(* IEC 61131-3 sources: codesys-ai-industrial-robot-control/plc/src/Tests, 11 files *)

(* ---- PRG_TestAlarms.st ---- *)
(*
    PRG_TestAlarms
    Purpose : Simulation test harness for FB_AlarmHandler (tests/plc/alarms.json).
    Inputs  : eId + xRaise / xRaiseEvent / xClear pulses, xAck, xReinit (each pulse resets itself).
*)
PROGRAM PRG_TestAlarms
VAR
    fbAlarms : FB_AlarmHandler;
    fbAlarmsInitial : FB_AlarmHandler;
    eId : E_AlarmId;
    xRaise : BOOL;
    xRaiseEvent : BOOL;
    xClear : BOOL;
    xAck : BOOL;
    xReinit : BOOL;
END_VAR

IF xReinit THEN
    xReinit := FALSE;
    fbAlarms := fbAlarmsInitial;
END_IF
IF xRaise THEN
    xRaise := FALSE;
    fbAlarms.Raise(eId);
END_IF
IF xRaiseEvent THEN
    xRaiseEvent := FALSE;
    fbAlarms.RaiseEvent(eId);
END_IF
IF xClear THEN
    xClear := FALSE;
    fbAlarms.Clear(eId);
END_IF
IF xAck THEN
    xAck := FALSE;
    fbAlarms.AcknowledgeAll();
END_IF
fbAlarms();

(* ---- PRG_TestCell.st ---- *)
(*
    PRG_TestCell
    Purpose : Simulation test harness for the whole cell in PRG_Main (tests/plc/cell.json).
              Simulates the vacuum switch, injects parts (PE1 pulse, then vision and decision
              messages for the captured part id) and can press the E-stop or lose the vacuum
              during a transfer. Can play the twin's bridge (heartbeat, joint feedback answering
              the current setpoint sample, twin active) and stall it. While active it plays an AI
              decision service (GVL_Bridge.xDecisionActive), reset when it is switched off.
    Inputs  : xActive; xInject (+ usiInjClass, eInjQuality); xEStopOnTransfer; xVacLostOnTransfer;
              xMark (J1 reference); xBridgeSim; xBridgeStall (heartbeat stops toggling);
              xBridgeStallOnTransfer
    Outputs : lrJ1Delta - J1 movement since xMark [deg]; lrAbortDelayMs - bridge stall -> Aborted
*)
PROGRAM PRG_TestCell
VAR
    xActive : BOOL;
    xWasActive : BOOL;
    xInject : BOOL;
    usiInjClass : USINT;
    eInjQuality : E_Quality := E_Quality.Ok;
    iInject : INT;
    tonPulse : TON;
    tonVac : TON;
    xEStopOnTransfer : BOOL;
    xVacLostOnTransfer : BOOL;
    xVacLost : BOOL;                    // latched until xVacLostOnTransfer is released
    xMark : BOOL;
    lrJ1Start : LREAL;
    lrJ1Delta : LREAL;
    xBridgeSim : BOOL;
    xBridgeStall : BOOL;
    xBridgeStallOnTransfer : BOOL;      // stall the bridge when the robot carries a part to its bin
    xStallTimed : BOOL;
    tStall : TIME;
    lrAbortDelayMs : LREAL;             // stall -> Aborted [ms]
END_VAR
VAR CONSTANT
    PE1_PULSE : TIME := T#250MS;
END_VAR

IF NOT xActive THEN
    IF xWasActive THEN                   // leave no fake decision service behind
        GVL_Bridge.xDecisionActive := FALSE;
        xWasActive := FALSE;
    END_IF
    RETURN;
END_IF
xWasActive := TRUE;
GVL_Bridge.xDecisionActive := TRUE;  // the harness injects AI decisions (eInjQuality)

IF xVacLostOnTransfer AND PRG_Main.fbCell.ePickStep = E_PickStep.MoveToBin THEN
    xVacLost := TRUE;
ELSIF NOT xVacLostOnTransfer THEN
    xVacLost := FALSE;
END_IF
tonVac(IN := GVL_Bridge.xVacuumOn, PT := T#100MS);
GVL_Bridge.xVacuumOk := tonVac.Q AND NOT xVacLost;

// the twin's bridge: feedback answers the current setpoint sample, heartbeat toggles
IF xBridgeStallOnTransfer AND NOT xBridgeStall AND PRG_Main.fbCell.ePickStep = E_PickStep.MoveToBin THEN
    xBridgeStall := TRUE;
    xStallTimed := FALSE;
    tStall := TIME();
END_IF
IF xBridgeStall AND NOT xStallTimed AND GVL_Bridge.eState = E_PackMLState.Aborted THEN
    xStallTimed := TRUE;
    lrAbortDelayMs := TIME_TO_LREAL(TIME() - tStall);
END_IF
IF xBridgeSim THEN
    GVL_Bridge.xTwinActive := TRUE;
    GVL_Bridge.aJointPosFb := GVL_Bridge.aJointPosSp;
    GVL_Bridge.udiFeedbackForSeq := GVL_Bridge.udiSetpointSeq;
    IF NOT xBridgeStall THEN
        GVL_Bridge.xHeartbeat := NOT GVL_Bridge.xHeartbeat;
        GVL_Bridge.udiFeedbackSeq := GVL_Bridge.udiFeedbackSeq + 1;
    END_IF
END_IF

CASE iInject OF
    0:
        IF xInject THEN
            xInject := FALSE;
            GVL_Bridge.xPE1 := TRUE;
            iInject := 1;
        END_IF
    1:
        tonPulse(IN := TRUE, PT := PE1_PULSE);
        IF tonPulse.Q THEN
            tonPulse(IN := FALSE);
            GVL_Bridge.xPE1 := FALSE;
            iInject := 2;
        END_IF
    2:
        GVL_Bridge.stVision.udiPartId := GVL_Bridge.stCapture.udiPartId;
        GVL_Bridge.stVision.xValid := TRUE;
        GVL_Bridge.stVision.usiClass := usiInjClass;
        GVL_Bridge.stVision.rConfidence := 0.9;
        GVL_Bridge.stVision.lrX := GVL_CellGeometry.PE1_X;
        GVL_Bridge.stVision.lrY := 0;
        GVL_Bridge.stVision.lrTheta := 0;
        GVL_Bridge.stVision.udiSeq := GVL_Bridge.stVision.udiSeq + 1;
        iInject := 3;
    3:
        GVL_Bridge.stDecision.udiPartId := GVL_Bridge.stVision.udiPartId;
        GVL_Bridge.stDecision.eQuality := eInjQuality;
        GVL_Bridge.stDecision.rQualityProb := 0.95;
        GVL_Bridge.stDecision.xIdentReliable := TRUE;
        GVL_Bridge.stDecision.udiSeq := GVL_Bridge.stDecision.udiSeq + 1;
        iInject := 0;
END_CASE

IF xEStopOnTransfer AND PRG_Main.fbCell.ePickStep = E_PickStep.MoveToBin THEN
    GVL_Bridge.xEStopOk := FALSE;
END_IF

IF xMark THEN
    xMark := FALSE;
    lrJ1Start := PRG_Main.fbCell.aActAcs[1];
END_IF
lrJ1Delta := PRG_Main.fbCell.aActAcs[1] - lrJ1Start;

(* ---- PRG_TestEquipment.st ---- *)
(*
    PRG_TestEquipment
    Purpose : Simulation test harness for the simple equipment FBs (tests/plc/equipment.json).
    Pulses  : write udiPulseMs and set xStartPulse - the harness drives fbPe.xRaw for exactly
              that long in PLC time (tool writes are too slow to time a short pulse).
*)
PROGRAM PRG_TestEquipment
VAR
    fbAlarms : FB_AlarmHandler;
    fbPe : FB_PhotoEye := (tDebounce := T#300MS);
    fbVac : FB_VacuumGripper;
    fbBin : FB_Bin := (eBin := E_Bin.TypeA);
    fbSafety : FB_SafetyMonitor;
    fbAlarmsInitial : FB_AlarmHandler;
    fbPeInitial : FB_PhotoEye := (tDebounce := T#300MS);
    fbVacInitial : FB_VacuumGripper;
    fbBinInitial : FB_Bin := (eBin := E_Bin.TypeA);
    fbSafetyInitial : FB_SafetyMonitor;
    xReinit : BOOL;
    uiPeRises : UINT;
    eVacError : E_AlarmId;
    udiPulseMs : UDINT;
    xStartPulse : BOOL;
    xPulseActive : BOOL;
    tonPulse : TON;
END_VAR

IF xReinit THEN
    xReinit := FALSE;
    fbAlarms := fbAlarmsInitial;
    fbPe := fbPeInitial;
    fbVac := fbVacInitial;
    fbBin := fbBinInitial;
    fbSafety := fbSafetyInitial;
    uiPeRises := 0;
    xPulseActive := FALSE;
END_IF
fbVac.itfAlarms := fbAlarms;
fbSafety.itfAlarms := fbAlarms;

IF xStartPulse THEN
    xStartPulse := FALSE;
    xPulseActive := TRUE;
END_IF
tonPulse(IN := xPulseActive, PT := TO_TIME(udiPulseMs));
IF tonPulse.Q THEN
    xPulseActive := FALSE;
END_IF
fbPe.xRaw := xPulseActive;

fbPe();
IF fbPe.xRising THEN
    uiPeRises := uiPeRises + 1;
END_IF
fbVac();
eVacError := fbVac.ErrorId;
fbBin();
fbSafety();
fbAlarms();

(* ---- PRG_TestJointMonitor.st ---- *)
(*
    PRG_TestJointMonitor
    Purpose : Simulation test harness for FB_JointMonitor (tests/plc/joint_monitor.json).
    Inputs  : xReinit; xAutoSeq - increment the feedback and setpoint sequences every cycle
              xRamp - J1 setpoint ramps by RAMP_STEP per cycle; iLag - feedback is the setpoint of
              iLag cycles earlier (and says so in udiFeedbackForSeq); xFreeze - feedback stands still;
              iTornSamples - that many cycles claim a sample iTornAge older (a torn OPC UA write,
              or a bridge hiccup when iTornAge exceeds the history)
    Outputs : lrRampSpeed - measured J1 setpoint speed [deg/s]
*)
PROGRAM PRG_TestJointMonitor
VAR
    fbMon : FB_JointMonitor;
    fbAlarms : FB_AlarmHandler;
    fbMonInitial : FB_JointMonitor;
    fbAlarmsInitial : FB_AlarmHandler;
    xReinit : BOOL;
    xAutoSeq : BOOL;
    xRamp : BOOL;
    xFreeze : BOOL;
    iLag : INT;
    udiSpSeq : UDINT;
    aSpHist : ARRAY[0..127] OF LREAL;
    xRampOld : BOOL;
    tRampStart : TIME;
    lrRampStart : LREAL;
    lrRampSpeed : LREAL;
    iTornSamples : INT;             // next cycles: feedback says it answers an older sample
    iTornAge : INT := 25;           // [samples]
END_VAR
VAR CONSTANT
    RAMP_STEP : LREAL := 1.0;       // [deg per cycle]
END_VAR

IF xReinit THEN
    xReinit := FALSE;
    xAutoSeq := FALSE;
    xRamp := FALSE;
    xFreeze := FALSE;
    iLag := 0;
    iTornSamples := 0;
    udiSpSeq := 0;
    fbMon := fbMonInitial;
    fbAlarms := fbAlarmsInitial;
END_IF
IF xAutoSeq THEN
    fbMon.udiFeedbackSeq := fbMon.udiFeedbackSeq + 1;
    udiSpSeq := udiSpSeq + 1;
END_IF
IF xRamp THEN
    IF NOT xRampOld THEN
        tRampStart := TIME();
        lrRampStart := fbMon.aSetpoint[1];
    END_IF
    fbMon.aSetpoint[1] := fbMon.aSetpoint[1] + RAMP_STEP;
    IF TIME() > tRampStart THEN
        lrRampSpeed := (fbMon.aSetpoint[1] - lrRampStart) * 1000.0 / TIME_TO_LREAL(TIME() - tRampStart);
    END_IF
END_IF
xRampOld := xRamp;
aSpHist[udiSpSeq MOD 128] := fbMon.aSetpoint[1];
fbMon.udiSetpointSeq := udiSpSeq;
IF udiSpSeq >= INT_TO_UDINT(iLag) THEN
    fbMon.udiFeedbackForSeq := udiSpSeq - INT_TO_UDINT(iLag);
    IF NOT xFreeze THEN
        fbMon.aFeedback[1] := aSpHist[fbMon.udiFeedbackForSeq MOD 128];
    END_IF
    IF iTornSamples > 0 AND fbMon.udiFeedbackForSeq >= INT_TO_UDINT(iTornAge) THEN
        fbMon.udiFeedbackForSeq := fbMon.udiFeedbackForSeq - INT_TO_UDINT(iTornAge);
        iTornSamples := iTornSamples - 1;
    END_IF
END_IF
fbMon.itfAlarms := fbAlarms;
fbMon();
fbAlarms();

(* ---- PRG_TestMotion.st ---- *)
(*
    PRG_TestMotion
    Purpose : Simulation test harness for FB_Robot and FB_Conveyor (tests/plc/motion.json).
    Inputs  : xActive - only then are the FBs called; xGo - start eCmd with the target chosen by
              iTargetSel (1 = home, 2 = current TCP - 50 mm in Z, 3 = home with J1 = 60 deg,
              4 = stProbe as written by the test)
    Outputs : xLastDone / xLastError of the last command, udiMoveMsLast / udiMoveMsPrev,
              xSlower (last move took > 1.5 x the previous one), lrZDelta
    Note    : SoftMotion FB instances are never re-initialised by assignment (corrupts them).
*)
PROGRAM PRG_TestMotion
VAR
    fbRobot : FB_Robot;
    fbConv : FB_Conveyor;
    fbAlarms : FB_AlarmHandler;
    xActive : BOOL;
    iTargetSel : INT;
    eCmd : E_RobotCmd;
    xGo : BOOL;
    iGoStep : INT;
    xLastDone : BOOL;
    xLastError : BOOL;
    tStart : TIME;
    udiMoveMsLast : UDINT;
    udiMoveMsPrev : UDINT;
    xSlower : BOOL;
    lrZStart : LREAL;
    lrZDelta : LREAL;
    stTarget : SMC_POS_REF;
    stProbe : SMC_POS_REF;
END_VAR

IF NOT xActive THEN
    RETURN;
END_IF
fbRobot.itfAlarms := fbAlarms;
fbConv.itfAlarms := fbAlarms;

IF xGo THEN
    xGo := FALSE;
    CASE iTargetSel OF
        1: stTarget := GVL_CellGeometry.HOME_ACS;
        2: stTarget := fbRobot.stActMcs;
           lrZStart := fbRobot.stActMcs.c.Z;
           stTarget.c.Z := lrZStart - 50;
        3: stTarget := GVL_CellGeometry.HOME_ACS;
           stTarget.a.a0 := 60;
        4: stTarget := stProbe;
    END_CASE
    fbRobot.stTarget := stTarget;
    fbRobot.eCmd := eCmd;
    fbRobot.xExecute := FALSE;     // a fresh rising edge, even if a command is running
    iGoStep := 1;
    xLastDone := FALSE;
    xLastError := FALSE;
ELSIF iGoStep = 1 THEN
    fbRobot.xExecute := TRUE;
    tStart := TIME();
    iGoStep := 2;
ELSIF iGoStep = 2 AND (fbRobot.xDone OR fbRobot.xError) THEN
    xLastDone := fbRobot.xDone;
    xLastError := fbRobot.xError;
    udiMoveMsPrev := udiMoveMsLast;
    udiMoveMsLast := TIME_TO_UDINT(TIME() - tStart);
    xSlower := udiMoveMsLast * 2 > udiMoveMsPrev * 3;
    fbRobot.xExecute := FALSE;
    iGoStep := 0;
END_IF

fbRobot(AxisGroup := AxisGroup_Robot);
fbConv(Axis := Axis_Conveyor);
fbAlarms();
IF iTargetSel = 2 THEN
    lrZDelta := fbRobot.stActMcs.c.Z - lrZStart;
END_IF

(* ---- PRG_TestMotionSmoke.st ---- *)
(*
    PRG_TestMotionSmoke
    Purpose : Simulation test harness - powers the robot axis group and makes one PTP move.
    Task    : TestTask (via PRG_Tests)
    Spec    : tests/plc/motion_smoke.json
*)
PROGRAM PRG_TestMotionSmoke
VAR
    fbPower : SMC_GroupPower;
    fbEnable : MC_GroupEnable;
    fbMove : MC_MoveDirectAbsolute := (CoordSystem := SMC_COORD_SYSTEM.ACS, VelFactor := 0.5);
    fbReadPos : MC_GroupReadActualPosition := (Enable := TRUE, CoordSystem := SMC_COORD_SYSTEM.ACS);
    xGo : BOOL;
    lrJ1 : LREAL;
    lrJ2 : LREAL;
    xMoveDone : BOOL;
    xMoveError : BOOL;
END_VAR

// Only commands the robot while the test runs, so other harnesses can use it.
IF xGo THEN
    fbPower(AxisGroup := AxisGroup_Robot, Enable := TRUE, bRegulatorOn := TRUE, bDriveStart := TRUE);
    fbEnable(AxisGroup := AxisGroup_Robot, Execute := fbPower.Status);
    fbMove.Position.a.a0 := 30;
    fbMove.Position.a.a1 := -20;
    fbMove.Position.a.a2 := 40;
    fbMove.Position.a.a3 := 0;
    fbMove.Position.a.a4 := 45;
    fbMove.Position.a.a5 := 0;
    fbMove(AxisGroup := AxisGroup_Robot, Execute := fbEnable.Done);
    fbReadPos(AxisGroup := AxisGroup_Robot);
    lrJ1 := fbReadPos.Position.a.a0;
    lrJ2 := fbReadPos.Position.a.a1;
    xMoveDone := fbMove.Done;
    xMoveError := fbMove.Error;
END_IF

(* ---- PRG_TestPackML.st ---- *)
(*
    PRG_TestPackML
    Purpose : Simulation test harness for FB_PackMLStateMachine (tests/plc/packml.json).
    Inputs  : xReinit - TRUE re-initialises the state machine, then resets itself.
*)
PROGRAM PRG_TestPackML
VAR
    fbSm : FB_PackMLStateMachine;
    fbSmInitial : FB_PackMLStateMachine;
    xReinit : BOOL;
END_VAR

IF xReinit THEN
    xReinit := FALSE;
    fbSm := fbSmInitial;
END_IF
fbSm();

(* ---- PRG_TestPick.st ---- *)
(*
    PRG_TestPick
    Purpose : Simulation test harness for FB_PickSequence (tests/plc/pick.json). Owns the robot,
              conveyor, gripper, tracker and alarms like the cell does, and simulates the vacuum
              switch (OK 100 ms after the valve opens).
    Inputs  : xActive, xBeltRun, xInject (+ usiInjClass, eInjQuality, lrInjX: one part with
              vision and decision; xInjInvalid: the vision message says "not seen"),
              xDropOnTransfer (vacuum lost during MoveToBin),
              xAbortOnLift (abort when the sequence reaches Lift), xResetSeq
    Outputs : xSawRecoverLift (latched: the recovery after an abort lifted first),
              lrGripZ (TCP height when the last grip started) [mm]
    Note    : SoftMotion FB instances are never re-initialised by assignment.
*)
PROGRAM PRG_TestPick
VAR
    fbRobot : FB_Robot;
    fbConv : FB_Conveyor;
    fbVac : FB_VacuumGripper;
    fbTracker : FB_PartTracker;
    fbAlarms : FB_AlarmHandler;
    fbSeq : FB_PickSequence;
    xActive : BOOL;
    xBeltRun : BOOL;
    xInject : BOOL;
    xInjInvalid : BOOL;
    usiInjClass : USINT;
    eInjQuality : E_Quality := E_Quality.Ok;
    lrInjX : LREAL := 1000;
    iInject : INT;
    xPE1 : BOOL;
    stVis : ST_VisionMsg;
    stDec : ST_DecisionMsg;
    xDropOnTransfer : BOOL;
    xAbortOnLift : BOOL;
    xResetSeq : BOOL;
    xVacLost : BOOL;
    tonVac : TON;
    xSawRecoverLift : BOOL;
    lrGripZ : LREAL;
    eLastStep : E_PickStep;
END_VAR

IF NOT xActive THEN
    RETURN;
END_IF
fbRobot.itfAlarms := fbAlarms;
fbConv.itfAlarms := fbAlarms;
fbVac.itfAlarms := fbAlarms;
fbTracker.itfAlarms := fbAlarms;
fbConv.xEnable := TRUE;
fbConv.lrVelocity := GVL_Params.lrBeltSpeed;
fbConv.xRun := xBeltRun;
fbRobot.xEnable := TRUE;

// One injected part: capture, then vision, then decision on consecutive cycles.
CASE iInject OF
    0:
        IF xInject THEN
            xInject := FALSE;
            xPE1 := TRUE;
            iInject := 1;
        END_IF
    1:
        xPE1 := FALSE;
        iInject := 2;
    2:
        stVis.udiSeq := stVis.udiSeq + 1;
        stVis.udiPartId := fbTracker.stCapture.udiPartId;
        stVis.xValid := NOT xInjInvalid;
        stVis.usiClass := usiInjClass;
        stVis.rConfidence := 0.9;
        stVis.lrX := lrInjX;
        stVis.lrY := 0;
        stVis.lrTheta := 0;
        iInject := 3;
    3:
        stDec.udiSeq := stDec.udiSeq + 1;
        stDec.udiPartId := stVis.udiPartId;
        stDec.eQuality := eInjQuality;
        stDec.rQualityProb := 0.95;
        stDec.xIdentReliable := TRUE;
        iInject := 0;
END_CASE

IF xDropOnTransfer AND fbSeq.eStep = E_PickStep.MoveToBin THEN
    xVacLost := TRUE;
END_IF
tonVac(IN := fbVac.xValveOn AND NOT xVacLost, PT := T#100MS);
fbVac.xVacuumOk := tonVac.Q;
IF xAbortOnLift AND fbSeq.eStep = E_PickStep.Lift THEN
    fbSeq.xAbort := TRUE;
END_IF
fbSeq.xReset := xResetSeq;
IF xResetSeq THEN
    xResetSeq := FALSE;
    xVacLost := FALSE;
    fbSeq.xAbort := FALSE;
    fbVac.Reset();
    fbAlarms.AcknowledgeAll();
END_IF

fbTracker(lrBeltPos := fbConv.lrPosition, xPE1Rising := xPE1, stVision := stVis, stDecision := stDec);
fbSeq(AxisGroup := AxisGroup_Robot, ConveyorAxis := Axis_Conveyor, Robot := fbRobot, Gripper := fbVac, Tracker := fbTracker);
fbVac();
fbRobot(AxisGroup := AxisGroup_Robot);
fbConv(Axis := Axis_Conveyor);
fbAlarms();
IF fbSeq.eStep = E_PickStep.RecoverLift THEN
    xSawRecoverLift := TRUE;
END_IF
IF fbSeq.eStep = E_PickStep.Grip AND eLastStep <> E_PickStep.Grip THEN
    lrGripZ := fbRobot.stActMcs.c.Z;
END_IF
eLastStep := fbSeq.eStep;

(* ---- PRG_Tests.st ---- *)
(*
    PRG_Tests
    Purpose : Calls every simulation test harness (TEST programs in this folder).
    Task    : TestTask, cyclic 10 ms
*)
PROGRAM PRG_Tests
VAR
END_VAR

PRG_TestMotionSmoke();
PRG_TestTypes();
PRG_TestPackML();
PRG_TestAlarms();
PRG_TestEquipment();
PRG_TestMotion();
PRG_TestJointMonitor();
PRG_TestTracking();
PRG_TestPick();
PRG_TestCell();

(* ---- PRG_TestTracking.st ---- *)
(*
    PRG_TestTracking
    Purpose : Simulation test harness for FB_PartTracker and F_SelectBin (tests/plc/tracking.json).
    Inputs  : lrBeltPos; xTriggerPE1 (one capture); uiFillCount (that many captures, one per cycle);
              stVisIn + xSendVision / xResendVision (same sequence number again);
              stDecIn + xSendDecision; udiQueryId - part to show in stRec; xAck; xClear;
              xNoDecisionLayer (no AI decision service)
    Outputs : uiCount, uiNext (next pickable index), stRec, xQueryFound
*)
PROGRAM PRG_TestTracking
VAR
    fbTracker : FB_PartTracker;
    fbAlarms : FB_AlarmHandler;
    fbTrackerInitial : FB_PartTracker;
    fbAlarmsInitial : FB_AlarmHandler;
    xReinit : BOOL;
    lrBeltPos : LREAL;
    xTriggerPE1 : BOOL;
    uiFillCount : UINT;
    stVisIn : ST_VisionMsg;
    stDecIn : ST_DecisionMsg;
    xSendVision : BOOL;
    xResendVision : BOOL;
    xSendDecision : BOOL;
    xAck : BOOL;
    xClear : BOOL;
    udiVisionSeq : UDINT;
    udiDecisionSeq : UDINT;
    udiQueryId : UDINT;
    uiQueryIdx : UINT;
    xQueryFound : BOOL;
    stRec : ST_PartRecord;
    uiCount : UINT;
    uiNext : UINT;
    xPE1Rising : BOOL;
    xNoDecisionLayer : BOOL;
END_VAR

IF xReinit THEN
    xReinit := FALSE;
    fbTracker := fbTrackerInitial;
    fbAlarms := fbAlarmsInitial;
    udiVisionSeq := 0;
    udiDecisionSeq := 0;
    uiFillCount := 0;
END_IF

xPE1Rising := xTriggerPE1 OR uiFillCount > 0;
xTriggerPE1 := FALSE;
IF uiFillCount > 0 THEN
    uiFillCount := uiFillCount - 1;
END_IF

IF xSendVision THEN
    xSendVision := FALSE;
    udiVisionSeq := udiVisionSeq + 1;
END_IF
IF xResendVision THEN
    xResendVision := FALSE;      // same sequence number: must be ignored
END_IF
stVisIn.udiSeq := udiVisionSeq;
IF xSendDecision THEN
    xSendDecision := FALSE;
    udiDecisionSeq := udiDecisionSeq + 1;
END_IF
stDecIn.udiSeq := udiDecisionSeq;
IF xAck THEN
    xAck := FALSE;
    fbAlarms.AcknowledgeAll();
END_IF
IF xClear THEN
    xClear := FALSE;
    fbTracker.Clear();
END_IF

fbTracker.itfAlarms := fbAlarms;
fbTracker(lrBeltPos := lrBeltPos, xPE1Rising := xPE1Rising, stVision := stVisIn, stDecision := stDecIn,
          xDecisionActive := NOT xNoDecisionLayer);
fbAlarms();

uiCount := fbTracker.Count;
uiNext := fbTracker.NextPickable(GVL_CellGeometry.PE2_X, GVL_CellGeometry.PICK_WINDOW_END_X);
uiQueryIdx := fbTracker.FindPart(udiQueryId);
xQueryFound := uiQueryIdx > 0;
IF xQueryFound THEN
    stRec := fbTracker.GetRecord(uiQueryIdx);
END_IF

(* ---- PRG_TestTypes.st ---- *)
(*
    PRG_TestTypes
    Purpose : Simulation test harness - exposes configuration values for tests/plc/types.json.
*)
PROGRAM PRG_TestTypes
VAR
    eClassBin0 : E_Bin;
    eFaultClass : E_AlarmClass;
    eWarnClass : E_AlarmClass;
    xLoopback : BOOL;
END_VAR

eClassBin0 := GVL_Params.aClassToBin[0];
eFaultClass := GVL_AlarmDefs.aDefs[E_AlarmId.EStop].eClass;
eWarnClass := GVL_AlarmDefs.aDefs[E_AlarmId.PartMissed].eClass;
xLoopback := GVL_Config.xFeedbackLoopback;
